(* IEC 61131-3 sources: SRCI_CLIENT_PLC/RobotLibrary/Library/POUs/General/MC_ReadServerLog/Structures, 4 files *)

(* ---- ReadServerLogOutCmd.st ---- *)
{attribute 'pack_mode' := '1'}
// -------------------------------------------------------------------------
//  SRCI Robot Library
// -------------------------------------------------------------------------
//
//  Object:      ReadServerLogOutCmd
//  Author:      Thorsten Brach
//  Date:        2026-10-23
//
//  Description:
//    Results of ReadServerLog (spec 6.2.6, table 6-120).
//
//  Copyright:
//    (C) 2026 Thorsten Brach. All rights reserved
//             Licensed under the MIT License.
//
//  Disclaimer:
//    This project is provided without any guarantee and can be used for
//    private and commercial purposes. Any use is at the user's
//    own risk and responsibility.
//
// -------------------------------------------------------------------------
TYPE ReadServerLogOutCmd :
STRUCT
  /// Total number of log lines in the requested log
  AvailableLogLines         : UDINT;
  /// Number of log lines in the requested log after the ContextFilter
  AvailableFilteredLogLines : UDINT;
  /// Number of log lines received and stored in LogFile (spec table 6-120: USINT)
  ReceivedLogLines          : UDINT;
  /// Received log lines compared to AvailableFilteredLogLines [%]
  Progress                  : REAL;
  /// The last log line of the requested log was transmitted
  EndOfLogReached           : BOOL;
  /// Number of the log line received last
  LogLine                   : UDINT;
END_STRUCT
END_TYPE

(* ---- ReadServerLogParCmd.st ---- *)
{attribute 'pack_mode' := '1'}
// -------------------------------------------------------------------------
//  SRCI Robot Library
// -------------------------------------------------------------------------
//
//  Object:      ReadServerLogParCmd
//  Author:      Thorsten Brach
//  Date:        2026-10-23
//
//  Description:
//    Parameters of ReadServerLog (spec 6.2.6, table 6-119).
//
//  Copyright:
//    (C) 2026 Thorsten Brach. All rights reserved
//             Licensed under the MIT License.
//
//  Disclaimer:
//    This project is provided without any guarantee and can be used for
//    private and commercial purposes. Any use is at the user's
//    own risk and responsibility.
//
// -------------------------------------------------------------------------
TYPE ReadServerLogParCmd :
STRUCT
  /// ID of the requested server log
  /// • -1 (default): latest server log
  /// •  0: oldest server log (SRCI SDK 1.1; spec table 6-119: 1)
  /// • >0: server log with this ID (OutCmd.ServerLogID of CreateServerLog)
  ServerLogID   : INT := -1;
  /// First log line of the requested log that is transferred to the PLC (1: log header)
  StartLine     : UDINT := 1;
  /// Only log lines of these contexts (spec table 6-118); all 0: no filter
  ContextFilter : ARRAY [0..9] OF USINT;
  /// Target of the log: 0 = output LogFile (default), 1 = export to a file (not supported)
  ExportMode    : USINT;
  /// File name of the export (ExportMode 1)
  ExportName    : STRING(20);
END_STRUCT
END_TYPE

(* ---- ReadServerLogRecvData.st ---- *)
{attribute 'pack_mode' := '1'}
// -------------------------------------------------------------------------
//  SRCI Robot Library
// -------------------------------------------------------------------------
//
//  Object:      ReadServerLogRecvData
//  Author:      Thorsten Brach
//  Date:        2026-10-23
//
//  Description:
//    Received CMD payload of ReadServerLog in the layout of SRCI SDK 1.1.2 (spec table 6-124:
//    only IsSplitLine, no EndOfLogReached / LogLine / Offset, 187 characters).
//
//  Copyright:
//    (C) 2026 Thorsten Brach. All rights reserved
//             Licensed under the MIT License.
//
//  Disclaimer:
//    This project is provided without any guarantee and can be used for
//    private and commercial purposes. Any use is at the user's
//    own risk and responsibility.
//
// -------------------------------------------------------------------------
TYPE ReadServerLogRecvData EXTENDS RspHeader :
STRUCT
  /// Total number of log lines in the requested log
  AvailableLogLines         : UDINT;
  /// Number of log lines after the ContextFilter
  AvailableFilteredLogLines : UDINT;
  /// Number of characters in LogContent
  LogContentLength          : USINT;
  /// Byte 13 Bit 0: LogContent starts a log line
  IsStartOfLine             : BOOL;
  /// Byte 13 Bit 1: LogContent ends a log line
  IsEndOfLine               : BOOL;
  /// Byte 13 Bit 2: the last log line was transmitted
  EndOfLogReached           : BOOL;
  /// Number of the transmitted log line
  LogLine                   : UDINT;
  /// Request counter of the command this response belongs to
  Offset                    : UDINT;
  /// Part of the log line (CSV)
  LogContent                : STRING(RobotLibraryConstants.SERVER_LOG_CONTENT_MAX);
END_STRUCT
END_TYPE

(* ---- ReadServerLogSendData.st ---- *)
{attribute 'pack_mode' := '1'}
// -------------------------------------------------------------------------
//  SRCI Robot Library
// -------------------------------------------------------------------------
//
//  Object:      ReadServerLogSendData
//  Author:      Thorsten Brach
//  Date:        2026-10-23
//
//  Description:
//    Sent CMD payload of ReadServerLog in the layout of SRCI SDK 1.1.2 (spec table 6-123
//    without Offset).
//
//  Copyright:
//    (C) 2026 Thorsten Brach. All rights reserved
//             Licensed under the MIT License.
//
//  Disclaimer:
//    This project is provided without any guarantee and can be used for
//    private and commercial purposes. Any use is at the user's
//    own risk and responsibility.
//
// -------------------------------------------------------------------------
TYPE ReadServerLogSendData EXTENDS CmdHeader :
STRUCT
  /// Byte 4 Bit 0: TRUE while log lines are transferred
  Enable        : BOOL;
  /// Reserve
  Reserve       : BYTE;
  /// ID of the requested server log (16#FFFF: latest, 0: oldest)
  ServerLogID   : UINT;
  /// First log line of the requested log
  StartLine     : UDINT;
  /// Request counter (SRCI SDK 1.1): every new value requests the next part of the log
  Offset        : UDINT;
  /// Only log lines of these contexts (spec table 6-118)
  ContextFilter : ARRAY [0..9] OF USINT;
END_STRUCT
END_TYPE
